Fanuc KAREL source: ka00079.KL

PROGRAM KA00079
%STACKSIZE=65535
%PRIORITY=65535
%NOLOCKGROUP
VAR
SRC : XYZWPREXT
DST : XYZWPREXT
BEGIN
SRC.X=1.0
DST=SRC
END KA00079
